// TIA Portal V20 export
// export: Created 2026-10-20T12:50:51.7738521Z, ExportSetting WithDefaults, DisplayName Totally Integrated Automation Portal, DisplayVersion V20 Update 6, DisplayName TIA Portal Openness, DisplayVersion V20 Update 6, DisplayName TIA Portal Version Control Interface, DisplayVersion V20 Update 6, DisplayName SINAMICS Startdrive Advanced, DisplayVersion V20 SP1, DisplayName SINAMICS Startdrive G130, G150, S120, S150, SINAMICS MV, G220, S200, S210, DisplayVersion V20 SP1, DisplayName SINAMICS Startdrive G110M, G120, G120C, G120D, G120P, G115D, DisplayVersion V20 SP1, DisplayName STEP 7 Professional, DisplayVersion V20 Update 6, DisplayName STEP 7 Safety, DisplayVersion V20 Update 2, DisplayName WinCC Basic/Comfort/Advanced, DisplayVersion V20 Update 6, DisplayName WinCC Unified, DisplayVersion V20 Update 6
FUNCTION_BLOCK "SICK Safe Entry Exit HW PLC V02"   // FB1000, F_FBD
TITLE = SICK Safe Entry Exit
AUTHOR : 2/29SD
FAMILY : S7-1500F
NAME : 9300351_02
VERSION : 2.0
// compiled for S7-1500F hardware controllers
// stored: IsIECCheckEnabled false, UDAEnableTagReadback false
   VAR_INPUT
      "########## BASIC_INPUTS ##########" : Bool := false;
      I_S_ESPE_Channel_1 : Bool := false;
      I_S_ESPE_Channel_2 : Bool := false;
      "I_S_PLC_request (MR)" : Bool := false;
      "I_S_Time_extension (TE)" : Bool := false;
      I_S_Reset : Bool := false;
      "I_S_Override hold-to-run-device" : Bool := false;
      I_S_first_logic_cycle : Bool := false;
      I_S_Disc_Time_MR_and_TE : Time := t#500ms;
      "########## MATERIAL_SELECTION_INPUTS ##########" : Bool := false;
      I_S_Material_selection_1 : Bool := false;
      I_S_Material_selection_2 : Bool := false;
      I_S_Material_selection_3 : Bool := false;
      I_S_Material_selection_4 : Bool := false;
      "########## MATERIAL_TOLERANCE_LENGTH in mm ##########" : Bool := false;
      "I_S_Material_tolerance_length_Material_1-4" : DInt := 100;
      "########## MAX_DISTANCE_MATERIAL_ESPE in mm ##########" : Bool := false;
      I_S_Max_distance_Material_to_ESPE : DInt := 0;
      "########## MATERIAL_LENGH_1-4 in mm ##########" : Bool := false;
      I_S_Material_length_Material_1 : DInt := 0;
      I_S_Material_length_Material_2 : DInt := 0;
      I_S_Material_length_Material_3 : DInt := 0;
      I_S_Material_length_Material_4 : DInt := 0;
      "########## MATERIAL_SPEED_1-4 in mm/s ##########" : Bool := false;
      I_S_Material_speed_Material_1 : DInt := 0;
      I_S_Material_speed_Material_2 : DInt := 0;
      I_S_Material_speed_Material_3 : DInt := 0;
      I_S_Material_speed_Material_4 : DInt := 0;
   END_VAR
   VAR_OUTPUT
      "########## BASIC_OUTPUTS ##########" : Bool := false;
      Q_Safety_release_1 : Bool := false;
      Q_Safety_release_2 : Bool;
      Q_SEE_Status : Bool := false;
      Q_Override_Status : Bool := false;
      Q_Reset_required : Bool := false;
      Q_Sequence_OK : Bool;
      "########## ERRORS ##########" : Bool := false;
      Error : Word := 0;
   END_VAR
   VAR
      "## BASIC SIGNALS ##" : Bool;
      ESPE : Bool;
      SEE_active : Bool;
      SEE_inactive : Bool;
      PLC_request : Bool;
      Time_extension : Bool;
      PLC_request_end : Bool;
      TE_signal_error : Bool;
      PLC_error : Bool;
      Timing_selection_error : Bool;
      Initiation_Error : Bool;
      SSE_aditional_release : Bool;
      Initiation : Bool;
      Termination : Bool;
      Termination_Seq_good : Bool;
      Override_status : Bool;
      Sequence_Signals_good : Bool;
      Material_1 : Bool;
      Material_2 : Bool;
      Material_3 : Bool;
      Material_4 : Bool;
      Min_time_good : Bool;
      Max_time_Error : Bool;
      TON_Tact_Lamps { S7_SetPoint := 'True'} : TON;
      TOF_Tact_Lamps { S7_SetPoint := 'True'} : TOF;
      Neg_Flag_Lamps : Bool;
      Blinking_tact : Bool;
      Always_0 : Bool := FALSE;
      Always_1 : Bool := TRUE;
      b_Sequence_Start : Bool;
      b_Sequence_OK : Bool;
      Sequence_OK { S7_SetPoint := 'True'} : TON;
      "## END BASIC SIGNALS ##" : Bool;
      "### CLOCK GENERATOR ###" : Bool;
      CLK_GEN_Edge_neg_1 : Bool;
      CLK_GEN_TON_Timer_1 { S7_SetPoint := 'True'} : TON;
      CLK_GEN_TOF_Timer_1 { S7_SetPoint := 'True'} : TOF;
      CLK_GEN_Tact : Bool;
      "### END CLOCK GENERATOR ###" : Bool;
      "### INITIATION ###" : Bool;
      INIT_HM_1 : Bool;
      INIT_HM_2 : Bool;
      INIT_HM_3 : Bool;
      INIT_Edge_neg_1 : Bool;
      "### END INITIATION ###" : Bool;
      "### MIN MAX TIME MONITORING ###" : Bool;
      MM_TIME_MONT_Fl_neg_1 : Bool;
      MM_TIME_MONT_TOF_Timer_1 { S7_SetPoint := 'True'} : TOF;
      MM_TIME_MONT_Int_timer_reset : Bool;
      MM_TIME_MONT_Counter_up_1 { S7_SetPoint := 'True'} : CTU;
      MM_TIME_MONT_Counter_up_2 { S7_SetPoint := 'True'} : CTU;
      MM_TIME_MONT_SEE_act_neg_edge : Bool;
      MM_TIME_MONT_Timer_reset : Bool;
      MM_TIME_MONT_TE_inactive : Bool;
      MM_TIME_MONT_TE_Timeout : Bool;
      MM_TIME_MONT_SEE_Timing_1 : Bool;
      MM_TIME_MONT_SEE_Timing_2 : Bool;
      MM_TIME_MONT_SEE_Timing_3 : Bool;
      MM_TIME_MONT_SEE_Timing_4 : Bool;
      "### END MIN MAX TIME MONITORING ###" : Bool;
      "### MULTIPLE STORE ###" : Bool;
      MUL_STORE_Edge_pos_1 : Bool;
      MUL_STORE_Save_Signal_1 : Bool;
      MUL_STORE_Save_Signal_2 : Bool;
      MUL_STORE_Save_Signal_3 : Bool;
      MUL_STORE_Save_Signal_4 : Bool;
      MUL_STORE_Save_Signal_5 : Bool;
      MUL_STORE_Save_Signal_6 : Bool;
      MUL_STORE_Save_Signal_7 : Bool;
      "### END MULTIPLE STORE ###" : Bool;
      "### OPERATION SELECTOR ###" : Bool;
      OP_SEL_Input_change : Bool;
      OP_SEL_Last_Cycle_Out_1 : Bool;
      OP_SEL_Last_Cycle_Out_2 : Bool;
      OP_SEL_Last_Cycle_Out_3 : Bool;
      OP_SEL_Last_Cycle_Out_4 : Bool;
      OP_SEL_Last_Cycle_Out_5 : Bool;
      OP_SEL_Last_Cycle_Out_6 : Bool;
      OP_SEL_Last_Cycle_Out_7 : Bool;
      OP_SEL_Last_Cycle_Out_8 : Bool;
      OP_SEL_HM_out_1 : Bool;
      OP_SEL_HM_out_2 : Bool;
      OP_SEL_HM_out_3 : Bool;
      OP_SEL_HM_out_4 : Bool;
      OP_SEL_HM_out_5 : Bool;
      OP_SEL_HM_out_6 : Bool;
      OP_SEL_HM_out_7 : Bool;
      OP_SEL_HM_out_8 : Bool;
      OP_SEL_TON_Timer_1 { S7_SetPoint := 'True'} : TON;
      OP_SEL_TON_Timer_2 { S7_SetPoint := 'True'} : TON;
      OP_SEL_Timing_1 : Bool;
      OP_SEL_Timing_2 : Bool;
      OP_SEL_Timing_3 : Bool;
      OP_SEL_Timing_4 : Bool;
      "### END OPERATION SELECTOR ###" : Bool;
      "### RESET1 ###" : Bool;
      RESET1_Edge_neg_1 : Bool;
      RESET1_M_Reset : Bool;
      RESET1_TON_TIMER_1 { S7_SetPoint := 'True'} : TON;
      RESET1_TON_TIMER_2 { S7_SetPoint := 'True'} : TON;
      RESET1_Release_OK : Bool;
      RESET1_Q : Bool;
      "### END RESET1 ###" : Bool;
      "### OVERRIDE ###" : Bool;
      OVR_TON_Timer_1 { S7_SetPoint := 'True'} : TON;
      OVR_Override_required : Bool;
      OVR_Override_status : Bool;
      OVR_Overriede_Clearance : Bool;
      "### END OVERRIDE ###" : Bool;
      "### RESET2 ###" : Bool;
      RESET2_Edge_neg_1 : Bool;
      RESET2_M_Reset : Bool;
      RESET2_TON_TIMER_1 { S7_SetPoint := 'True'} : TON;
      RESET2_TON_TIMER_2 { S7_SetPoint := 'True'} : TON;
      RESET2_Release_OK : Bool;
      "### END RESET2 ###" : Bool;
      "### TERMINATION ###" : Bool;
      TERM_Edge_neg_1 : Bool;
      TERM_Edge_pos_1 : Bool;
      TERM_HM_1 : Bool;
      TERM_TOF_Timer_1 { S7_SetPoint := 'True'} : TOF;
      "### END TERMINATION ###" : Bool;
      "### MIN_MAX_TIMER_RESET ###" : Bool;
      MIN_MAX_TIME_TON_Timer_Reset { S7_SetPoint := 'True'} : TON;
      "### END_MIN_MAX_TIMER_RESET ###" : Bool;
      "###MIN TIME  ###" : Bool;
      MIN_TIME_1_Timer_save : Time;
      MIN_TIME_1_Timer_1st_stop : Bool := FALSE;
      MIN_TIME_1_Edge_neg_1 : Bool;
      MIN_TIME_1_TON_Timer_1 { S7_SetPoint := 'True'} : TON;
      MIN_TIME_1_Q : Bool;
      MIN_TIME_2_Timer_save : Time;
      MIN_TIME_2_Timer_1st_stop : Bool := FALSE;
      MIN_TIME_2_Edge_neg : Bool;
      MIN_TIME_2_TON_Timer { S7_SetPoint := 'True'} : TON;
      MIN_TIME_2_Q : Bool;
      MIN_TIME_3_Timer_save : Time;
      MIN_TIME_3_Timer_1st_stop : Bool;
      MIN_TIME_3_Edge_neg : Bool;
      MIN_TIME_3_TON_Timer { S7_SetPoint := 'True'} : TON;
      MIN_TIME_3_Q : Bool;
      MIN_TIME_4_Timer_save : Time;
      MIN_TIME_4_Timer_1st_stop : Bool;
      MIN_TIME_4_Edge_neg : Bool;
      MIN_TIME_4_TON_Timer { S7_SetPoint := 'True'} : TON;
      MIN_TIME_4_Q : Bool;
      "###END MIN TIME ###" : Bool;
      "###MAX TIME  ###" : Bool;
      MAX_TIME_1_Timer_save : Time;
      MAX_TIME_1_Timer_1st_stop : Bool;
      MAX_TIME_1_Edge_neg : Bool;
      MAX_TIME_1_TON_Timer { S7_SetPoint := 'True'} : TON;
      MAX_TIME_1_Q : Bool;
      MAX_TIME_2_Timer_save : Time;
      MAX_TIME_2_Timer_1st_stop : Bool;
      MAX_TIME_2_Edge_neg : Bool;
      MAX_TIME_2_TON_Timer { S7_SetPoint := 'True'} : TON;
      MAX_TIME_2_Q : Bool;
      MAX_TIME_3_Timer_save : Time;
      MAX_TIME_3_Timer_1st_stop : Bool;
      MAX_TIME_3_Edge_neg : Bool;
      MAX_TIME_3_TON_Timer { S7_SetPoint := 'True'} : TON;
      MAX_TIME_3_Q : Bool;
      MAX_TIME_4_Timer_save : Time;
      MAX_TIME_4_Timer_1st_stop : Bool;
      MAX_TIME_4_Edge_neg : Bool;
      MAX_TIME_4_TON_Timer { S7_SetPoint := 'True'} : TON;
      MAX_TIME_4_Q : Bool;
      "###END MAX TIME  ###" : Bool;
      "### DISC CONTROL 1 ###" : Bool;
      DISC_1_b_Input_A : Bool;
      DISC_1_b_Input_B : Bool;
      DISC_1_Fl_pos_1 : Bool;
      DISC_1_Fl_neg_1 : Bool;
      DISC_1_Fl_neg_2 : Bool;
      DISC_1_Startbit : Bool;
      DISC_1_Stopbit : Bool;
      DISC_1_M_Release : Bool;
      DISC_1_M_AND_Mode_active : Bool;
      DISC_1_TON_Timer_1 { S7_SetPoint := 'True'} : TON;
      DISC_1_TON_Timer_2 { S7_SetPoint := 'True'} : TON;
      DISC_1_TON_Timer_3 { S7_SetPoint := 'True'} : TON;
      DISC_1_TOF_Timer_1 { S7_SetPoint := 'True'} : TOF;
      DISC_1_TOF_Timer_2 { S7_SetPoint := 'True'} : TOF;
      DISC_1_Q : Bool;
      DISC_1_Error : Bool;
      DISC_1_Error_Discrepancy_1 : Bool;
      DISC_1_Error_Discrepancy_2 : Bool;
      "### END DISC CONTROL 1 ###" : Bool;
      "### DISC CONTROL 2 ###" : Bool;
      DISC_2_b_Input_A : Bool;
      DISC_2_b_Input_B : Bool;
      DISC_2_Fl_pos_1 : Bool;
      DISC_2_Fl_neg_1 : Bool;
      DISC_2_Fl_neg_2 : Bool;
      DISC_2_Startbit : Bool;
      DISC_2_Stopbit : Bool;
      DISC_2_M_Release : Bool;
      DISC_2_M_AND_Mode_active : Bool;
      DISC_2_TON_Timer_1 { S7_SetPoint := 'True'} : TON;
      DISC_2_TON_Timer_2 { S7_SetPoint := 'True'} : TON;
      DISC_2_TON_Timer_3 { S7_SetPoint := 'True'} : TON;
      DISC_2_TOF_Timer_1 { S7_SetPoint := 'True'} : TOF;
      DISC_2_TOF_Timer_2 { S7_SetPoint := 'True'} : TOF;
      DISC_2_Q : Bool;
      DISC_2_Error : Bool;
      DISC_2_Error_Discrepancy_2 : Bool;
      DISC_2_Error_Discrepancy_1 : Bool;
      "### END DISC CONTROL 2 ###" : Bool;
      "### PLC SIG MONITORING ###" : Bool;
      PLC_SIG_MON_Edge_pos_1 : Bool;
      PLC_SIG_MON_Edge_neg_1 : Bool;
      PLC_SIG_MON_Edge_neg_2 : Bool;
      PLC_SIG_MON_HM_1 : Bool;
      PLC_SIG_MON_Int_muting_request : Bool;
      PLC_SIG_MON_Int_time_extension : Bool;
      PLC_SIG_MON_Discrepancy_control_Q : Bool;
      PLC_SIG_MON_Error_discrepancy_control_1 : Bool;
      PLC_SIG_MON_TON_Timer_1 { S7_SetPoint := 'True'} : TON;
      "### END PLC SIG MONITORING ###" : Bool;
      "### SSE #####" : Bool;
      SSE_Int_Enable : Bool;
      SSE_Int_Muting_active : Bool;
      SSE_Int_Safe_condition : Bool;
      "### END SSE #####" : Bool;
      "### SEQUENCE MONITORING ###" : Bool;
      SEQ_MON_TOF_Timer_1 { S7_SetPoint := 'True'} : TOF;
      SEQ_MON_TOF_Timer_2 { S7_SetPoint := 'True'} : TOF;
      SEQ_MON_TOF_Timer_3 { S7_SetPoint := 'True'} : TOF;
      SEQ_MON_TOF_Timer_4 { S7_SetPoint := 'True'} : TOF;
      SEQ_MON_TON_Timer_5 { S7_SetPoint := 'True'} : TON;
      SEQ_MON_TON_Timer_6 { S7_SetPoint := 'True'} : TON;
      SEQ_MON_TON_Timer_7 { S7_SetPoint := 'True'} : TON;
      SEQ_MON_TON_Timer_8 { S7_SetPoint := 'True'} : TON;
      SEQ_MON_TON_Timer_9 { S7_SetPoint := 'True'} : TON;
      SEQ_MON_TON_Timer_10 { S7_SetPoint := 'True'} : TON;
      SEQ_MON_TON_Timer_11 { S7_SetPoint := 'True'} : TON;
      SEQ_MON_TON_Timer_12 { S7_SetPoint := 'True'} : TON;
      SEQ_MON_Edge_PLC_request : Bool;
      SEQ_MON_Edge_pos_1 : Bool;
      SEQ_MON_Error_PLC_Req : Bool;
      SEQ_MON_HM_PLC_request : Bool;
      "### END SEQUENCE MONITORING ###" : Bool;
      "### ERROR HANDLING ###" : Bool;
      ERR_Handling_INT : Int;
      ERR_Handling_Neg_Flag : Bool;
      ERR_Signal_monitoring_MR_TE : Bool;
      ERR_Signal_monitoring_MR_TE_direct : Bool;
      HM_Sequenz_MR_TE_1 : Bool;
      HM_Sequenz_MR_TE_2 : Bool;
      HM_Sequenz_MR_TE_OK : Bool;
      ERR_Flag_Pos : Bool;
      ERR_FL_Neg : Bool;
      TON_Timer_Err_direct { S7_SetPoint := 'True'} : TON;
      "Create Error Termination Sequence" : Bool;
      "Create Error Min time" : Bool;
      "Create Error Max time" : Bool;
      "Create Error Timing selection" : Bool;
      "Create Error PLC Signal" : Bool;
      "Create Error TE Signal" : Bool;
      "Create Error Discrepancy MR TE" : Bool;
      "Create Error Discrepancy ESPE" : Bool;
      "Create Error calculation zero" : Bool;
      "Create Error Signal monitoring MR TE" : Bool;
      "Create Error Max. Dist ESPE" : Bool;
      "Create Error Monitoring Max. Muting" : Bool;
      "Create Error Max. INIT Time" : Bool;
      "Create Error Initiation sequence" : Bool;
      "Create Error min time less 500mm" : Bool;
      Reset_bit : Bool;
      "### END ERROR HANDLING ###" : Bool;
   END_VAR
BEGIN
END_FUNCTION_BLOCK
